(* IEC 61131-3 sources: llm-plc-st-eval/data/processed_v2_primera/claude-sonnet-4-6/I5/zero_shot, 3 files *)

(* ---- ejec_1.st ---- *)
FUNCTION_BLOCK FB_Clasificadora
VAR_INPUT
    sensorPresencia : BOOL; (* Sensor de paso de pieza *)
    sensorAltura    : BOOL; (* TRUE = pieza alta *)
END_VAR

VAR_OUTPUT
    banda   : BOOL; (* Banda transportadora activa *)
    piston  : BOOL; (* Desviador activo *)
    nAltas  : INT;  (* Contador de piezas altas *)
    nBajas  : INT;  (* Contador de piezas bajas *)
END_VAR

VAR
    tRetardo    : TON; (* Temporizador retardo 2 s hasta el desviador *)
    tPiston     : TON; (* Temporizador duración del pistón 1 s *)
    rPresencia  : R_TRIG; (* Flanco ascendente del sensor de presencia *)
    bPiezaAlta  : BOOL;   (* Indica que la pieza detectada es alta *)
    bEsperando  : BOOL;   (* TRUE mientras se espera el retardo *)
END_VAR

(* ── Banda siempre activa ─────────────────────────────────────── *)
banda := TRUE;

(* ── Detección de flanco en sensorPresencia ───────────────────── *)
rPresencia(CLK := sensorPresencia);

IF rPresencia.Q THEN
    (* Nueva pieza detectada *)
    IF sensorAltura THEN
        (* Pieza alta: registrar y armar retardo *)
        nAltas     := nAltas + 1;
        bPiezaAlta := TRUE;
        bEsperando := TRUE;
    ELSE
        (* Pieza baja: solo contar *)
        nBajas := nBajas + 1;
    END_IF;
END_IF;

(* ── Retardo de 2 s (pieza viaja hasta el desviador) ─────────── *)
tRetardo(IN := bEsperando, PT := T#2S);

IF tRetardo.Q THEN
    (* Han pasado 2 s: activar pistón y detener retardo *)
    bEsperando := FALSE;
    tRetardo(IN := FALSE);  (* Reset del temporizador de retardo *)
    bPiezaAlta := TRUE;     (* Señal para arrancar temporizador pistón *)
END_IF;

(* ── Activación del pistón durante 1 s ───────────────────────── *)
tPiston(IN := tRetardo.Q OR tPiston.Q AND NOT tPiston.ET = T#1S, PT := T#1S);
(* Nota: se usa el flanco de salida de tRetardo para arrancar tPiston *)
tPiston(IN := (tRetardo.Q), PT := T#1S);

piston := tPiston.Q OR (tRetardo.Q);

(* ── Salida limpia del pistón ─────────────────────────────────── *)
(* tPiston corre mientras su entrada IN sea TRUE;
   se mantiene TRUE hasta que ET alcance PT (1 s) *)
IF tPiston.ET >= T#1S THEN
    tPiston(IN := FALSE);   (* Reset del temporizador del pistón *)
    piston := FALSE;
END_IF;

END_FUNCTION_BLOCK

(* ---- ejec_2.st ---- *)
FUNCTION_BLOCK FB_Clasificadora
VAR_INPUT
    sensorPresencia : BOOL; (* Sensor de paso de pieza *)
    sensorAltura    : BOOL; (* TRUE = pieza alta *)
END_VAR

VAR_OUTPUT
    banda   : BOOL; (* Salida banda transportadora *)
    piston  : BOOL; (* Salida pistón desviador *)
    nAltas  : INT;  (* Contador de piezas altas *)
    nBajas  : INT;  (* Contador de piezas bajas *)
END_VAR

VAR
    tRetardo    : TON; (* Temporizador retardo 2 s hasta el desviador *)
    tPiston     : TON; (* Temporizador duración del pistón 1 s *)
    rPresencia  : R_TRIG; (* Flanco ascendente del sensor de presencia *)
    bPiezaAlta  : BOOL;   (* Indica que la pieza detectada es alta *)
    bContado    : BOOL;   (* Evita contar la misma pieza más de una vez *)
END_VAR

(* ------------------------------------------------------------------ *)
(* 1. La banda funciona siempre                                        *)
(* ------------------------------------------------------------------ *)
banda := TRUE;

(* ------------------------------------------------------------------ *)
(* 2. Detectar flanco ascendente del sensor de presencia              *)
(* ------------------------------------------------------------------ *)
rPresencia(CLK := sensorPresencia);

IF rPresencia.Q THEN
    (* Capturar si la pieza es alta en el momento de la detección *)
    bPiezaAlta := sensorAltura;
    bContado   := FALSE;

    IF bPiezaAlta THEN
        (* Arrancar el retardo de 2 s antes de activar el pistón *)
        tRetardo.IN := FALSE; (* Reset previo para reiniciar el temporizador *)
    END_IF;
END_IF;

(* ------------------------------------------------------------------ *)
(* 3. Gestión del retardo (2 s) y del pistón (1 s) para piezas altas *)
(* ------------------------------------------------------------------ *)
(* Activar el temporizador de retardo mientras haya pieza alta pendiente
   y el pistón aún no haya terminado su ciclo                         *)
tRetardo(IN := bPiezaAlta AND NOT tRetardo.Q,
         PT := T#2S);

(* Cuando el retardo termina, activar el temporizador del pistón *)
tPiston(IN := tRetardo.Q AND NOT tPiston.Q,
        PT := T#1S);

(* Salida del pistón activa durante el segundo de accionamiento *)
piston := tRetardo.Q AND NOT tPiston.Q;

(* ------------------------------------------------------------------ *)
(* 4. Conteo de piezas y limpieza de estado al finalizar el ciclo     *)
(* ------------------------------------------------------------------ *)
IF bPiezaAlta AND tPiston.Q AND NOT bContado THEN
    (* Ciclo completo de pieza alta: retardo + pistón terminados *)
    nAltas   := nAltas + 1;
    bContado := TRUE;

    (* Resetear temporizadores y bandera para el siguiente ciclo *)
    tRetardo.IN := FALSE;
    tPiston.IN  := FALSE;
    bPiezaAlta  := FALSE;
END_IF;

IF NOT bPiezaAlta AND rPresencia.Q THEN
    (* Pieza baja: contar en el mismo ciclo de detección *)
    nBajas := nBajas + 1;
END_IF;

END_FUNCTION_BLOCK

(* ---- ejec_3.st ---- *)
FUNCTION_BLOCK FB_Clasificadora
VAR_INPUT
    sensorPresencia : BOOL; (* Sensor de paso de pieza *)
    sensorAltura    : BOOL; (* TRUE = pieza alta *)
END_VAR

VAR_OUTPUT
    banda   : BOOL; (* Banda transportadora activa *)
    piston  : BOOL; (* Desviador activo *)
    nAltas  : INT;  (* Contador de piezas altas *)
    nBajas  : INT;  (* Contador de piezas bajas *)
END_VAR

VAR
    tRetardo    : TON; (* Temporizador retardo 2 s hasta el desviador *)
    tPiston     : TON; (* Temporizador duración del pistón 1 s *)
    rPresencia  : R_TRIG; (* Flanco ascendente del sensor de presencia *)
    piezaAlta   : BOOL;   (* Indica que la pieza detectada es alta *)
END_VAR

(* ── Banda siempre activa ─────────────────────────────────────── *)
banda := TRUE;

(* ── Detección de flanco en sensorPresencia ───────────────────── *)
rPresencia(CLK := sensorPresencia);

IF rPresencia.Q THEN
    (* Nueva pieza detectada: registrar su tipo y arrancar retardo *)
    piezaAlta := sensorAltura;

    IF piezaAlta THEN
        nAltas := nAltas + 1; (* Contar pieza alta *)
    ELSE
        nBajas := nBajas + 1; (* Contar pieza baja *)
    END_IF;

    (* Reiniciar temporizadores para esta pieza *)
    tRetardo(IN := FALSE, PT := T#2S);
    tPiston (IN := FALSE, PT := T#1S);
END_IF;

(* ── Retardo de 2 s: tiempo de tránsito hasta el desviador ───── *)
IF piezaAlta THEN
    tRetardo(IN := TRUE, PT := T#2S);
ELSE
    tRetardo(IN := FALSE, PT := T#2S);
END_IF;

(* ── Activar pistón durante 1 s al cumplirse el retardo ─────── *)
IF tRetardo.Q THEN
    tPiston(IN := TRUE, PT := T#1S); (* Arrancar temporizador pistón *)
END_IF;

IF tPiston.Q THEN
    (* Tiempo de pistón cumplido: desactivar todo *)
    tPiston (IN := FALSE, PT := T#1S);
    tRetardo(IN := FALSE, PT := T#2S);
    piezaAlta := FALSE;
END_IF;

(* ── Salida pistón activa mientras tPiston está contando ─────── *)
piston := tPiston.IN AND NOT tPiston.Q;

END_FUNCTION_BLOCK
